(* IEC 61131-3 sources: kns-pump-station/tests/POUs/Station/FB_Ventilation_Test, 6 files *)

(* ---- FireInterlocksAndStops.method.decl.st ---- *)
// 04 §17, PMI-38: пожар — В1 стоп и блокировка V1_ILK_FIRE при любых условиях
METHOD PRIVATE FireInterlocksAndStops
VAR
    fbDut  : FB_Ventilation;            // ФБ под тестом
    fbTime : PL.FB_FakeTime;            // подменное время, старт 1 ч
    stCfg  : ST_StationCfg;             // уставки по умолчанию: выбег 10 мин
END_VAR

(* ---- OverrunAfterConditionsClear.method.decl.st ---- *)
// 04 §17, PMI-38: условия сняты — В1 работает ещё tV1Overrun = 10 мин, затем стоп
METHOD PRIVATE OverrunAfterConditionsClear
VAR
    fbDut  : FB_Ventilation;            // ФБ под тестом
    fbTime : PL.FB_FakeTime;            // подменное время, старт 1 ч
    stCfg  : ST_StationCfg;             // уставки по умолчанию: выбег 10 мин
    uiStep : UINT;                      // шаг 1 с
END_VAR

(* ---- OverrunAfterConditionsClear.method.impl.st ---- *)
coUnit.TEST('Ventilation_OverrunAfterConditionsClear_A17_PMI38');

fbDut(xDoorOpen := TRUE, itfTime := fbTime, stCfg := stCfg);
fbTime.Advance(tStep := T#1S);
fbDut(xDoorOpen := FALSE, itfTime := fbTime, stCfg := stCfg);
FOR uiStep := 1 TO 599 DO
    fbTime.Advance(tStep := T#1S);
    fbDut(itfTime := fbTime, stCfg := stCfg);
END_FOR
AssertTrue(Condition := fbDut.xRun, Message := 'overrun at 9 min 59 s');
fbTime.Advance(tStep := T#1S);
fbDut(itfTime := fbTime, stCfg := stCfg);
AssertFalse(Condition := fbDut.xRun, Message := 'stop at 10 min');

coUnit.TEST_FINISHED();

(* ---- RunsOnGasDoorTemp.method.decl.st ---- *)
// 04 §17, PMI-38: В1 работает при газе выше H, открытой двери, температуре выше H
METHOD PRIVATE RunsOnGasDoorTemp
VAR
    fbDut  : FB_Ventilation;            // ФБ под тестом
    fbTime : PL.FB_FakeTime;            // подменное время, старт 1 ч
    stCfg  : ST_StationCfg;             // уставки по умолчанию: выбег 10 мин
    fbDut2 : FB_Ventilation;           // дверь
    fbDut3 : FB_Ventilation;           // температура
END_VAR

(* ---- TimeBackwardsRestartsOverrun.method.decl.st ---- *)
// Время назад — выбег tV1Overrun отсчитывается заново (вентилятор работает дольше, а не останавливается раньше)
METHOD PRIVATE TimeBackwardsRestartsOverrun
VAR
    fbDut  : FB_Ventilation;            // ФБ под тестом
    fbTime : PL.FB_FakeTime;            // подменное время, старт 1 ч
    stCfg  : ST_StationCfg;             // уставки по умолчанию: выбег 10 мин
    uiStep : UINT;                      // шаг 1 с
END_VAR

(* ---- TimeBackwardsRestartsOverrun.method.impl.st ---- *)
coUnit.TEST('Ventilation_TimeBackwardsRestartsOverrun_A17');

fbDut(xDoorOpen := TRUE, itfTime := fbTime, stCfg := stCfg);
fbTime.Advance(tStep := T#1S);
fbDut(xDoorOpen := FALSE, itfTime := fbTime, stCfg := stCfg);
FOR uiStep := 1 TO 100 DO
    fbTime.Advance(tStep := T#1S);
    fbDut(itfTime := fbTime, stCfg := stCfg);
END_FOR
fbTime.SetNow(ltValue := LTIME#59M);
FOR uiStep := 1 TO 600 DO
    fbTime.Advance(tStep := T#1S);
    fbDut(itfTime := fbTime, stCfg := stCfg);
END_FOR
AssertTrue(Condition := fbDut.xRun, Message := 'overrun restarted after time jump');
fbTime.Advance(tStep := T#1S);
fbDut(itfTime := fbTime, stCfg := stCfg);
AssertFalse(Condition := fbDut.xRun, Message := 'stop after full overrun');

coUnit.TEST_FINISHED();
